Fanuc KAREL source: ka00144.KL

-- PROVISIONAL review KL for V940-1; original PC SHA256 221dc29e801ddfb958c89b92d92a72b5b3428f65c97f0c2e4c399efada2391eb
-- Incomplete behavior may be omitted. Consult companion uncertainty JSON. Do not deploy.
PROGRAM KA00144
%NOLOCKGROUP
-- UNRESOLVED_DECL SRC type=002017
-- UNRESOLVED_DECL DST type=002017
BEGIN
  -- V9_ZERO_TABLE_METADATA_HINT layout=0001; no indexed target words; source/name/runtime held
  -- UNRESOLVED_PC offsets 5-19; opcodes 2E,22,9D,33,B4
  -- UNRESOLVED_PC offsets 24-42; opcodes 22,9D,33,B3,22,9D,33,B4
  -- UNRESOLVED_PC offsets 47-51; opcodes 7F
END KA00144
